TYPE ST_PLCTOLEISTER :
STRUCT
	arbyOutput				:ARRAY[0..63] OF BYTE;
END_STRUCT
END_TYPE

(* stored: Version 1.1.0.1, ProductVersion 3.1.4024.15
   DUT ST_PLCTOLEISTER: Id {5a5ee05e-f634-4790-8122-dda71dc82aef} *)
